Fanuc KAREL source: KT00680.KL

PROGRAM KT00680
%NOLOCKGROUP
VAR
  P1: JOINTPOS
  P2: JOINTPOS
  OUT: REAL
BEGIN
  OUT = NOT P1
END KT00680
